(* PLC project Vn_fanout_into_box, Beckhoff Automation GmbH TwinCAT PLC Control 3.5.13.21 *)
(* stored: creationDateTime 1970-01-01T00:00:00 *)

PROGRAM Vn_fanout_into_box
  VAR  (* added by the conversion: wires and edge detectors of the diagram *)
    _AND10000000003_OUT : BOOL;
  END_VAR

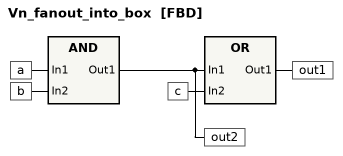
(* FBD diagram, written out as Structured Text *)
_AND10000000003_OUT := a AND b;
out1 := _AND10000000003_OUT OR c;
out2 := _AND10000000003_OUT;
END_PROGRAM
